Fanuc KAREL source: kd00049.KL

-- PROVISIONAL review KL for V1013-1; original PC SHA256 a1cd803d81ce8b2f60a28f7ad37f3ed6e8bad5934bec1b73c483a0b382cfc6f2
-- Incomplete behavior may be omitted. Consult companion uncertainty JSON. Do not deploy.
PROGRAM KD00049
%NOLOCKGROUP
VAR
  I : INTEGER
  J : INTEGER
  B : BOOLEAN
  R : REAL
  S : STRING[80]
BEGIN
  -- UNRESOLVED_PC offsets 5-18; opcodes 01,2E,0A,82,0B
  -- UNRESOLVED_PC offsets 23-27; opcodes 7F
END KD00049
